// TIA Portal V21 export
// export: Created 2026-11-10T19:12:20.8340068Z, ExportSetting WithDefaults, DisplayName Totally Integrated Automation Portal, DisplayVersion V21 Update 3, DisplayName STEP 7 Professional, DisplayVersion V21 Update 3, DisplayName STEP 7 Safety, DisplayVersion V21, DisplayName Tech WebApplication, DisplayVersion V21, DisplayName WinCC Basic/Comfort/Advanced, DisplayVersion V21 Update 3, DisplayName WinCC Unified, DisplayVersion V21 Update 3
DATA_BLOCK "DBsCONT_C"   // DB31
// stored: AutoNumber true, DBAccessibleFromOPCUA true, DBAccessibleFromWebserver true, InstanceOfName CONT_C, OfSystemLibElement CONT_C, OfSystemLibVersion 1.1
CONT_C   // technology object, version 1.1
   // VAR_INPUT
   //    COM_RST : Bool;
   //    MAN_ON : Bool;
   //    PVPER_ON : Bool;
   //    P_SEL : Bool;
   //    I_SEL : Bool;
   //    INT_HOLD : Bool;
   //    I_ITL_ON : Bool;
   //    D_SEL : Bool;
   //    CYCLE : Time;
   //    SP_INT : Real;
   //    PV_IN : Real;
   //    PV_PER : Word;
   //    MAN : Real;
   //    GAIN : Real;
   //    TI : Time;
   //    TD : Time;
   //    TM_LAG : Time;
   //    DEADB_W : Real;
   //    LMN_HLM : Real;
   //    LMN_LLM : Real;
   //    PV_FAC : Real;
   //    PV_OFF : Real;
   //    LMN_FAC : Real;
   //    LMN_OFF : Real;
   //    I_ITLVAL : Real;
   //    DISV : Real;
   // END_VAR
   // VAR_OUTPUT
   //    LMN : Real;
   //    LMN_PER : Word;
   //    QLMN_HLM : Bool;
   //    QLMN_LLM : Bool;
   //    LMN_P : Real;
   //    LMN_I : Real;
   //    LMN_D : Real;
   //    PV : Real;
   //    ER : Real;
   // END_VAR
   // VAR RETAIN
   //    sInvAlt : Real;
   //    sIanteilAlt : Real;
   //    sRestInt : Real;
   //    sRestDif : Real;
   //    sRueck : Real;
   //    sLmn : Real;
   //    sbArwHLmOn : Bool;
   //    sbArwLLmOn : Bool;
   //    sbILimOn : Bool;
   // END_VAR
BEGIN
END_DATA_BLOCK
